(* IEC 61131-3 sources: avi-aoi-management/scripts/ai-eval/ngau-nhien/kho/st-ud7-van-hai-cuon/khung/src, 2 files *)

(* ---- ViTriVan.st ---- *)
FUNCTION ViTriVan : INT
VAR_INPUT
    CT_MO : BOOL;
    CT_DONG : BOOL;
END_VAR
    (* TODO: cài đặt theo đề bài *)
    ViTriVan := -1;
END_FUNCTION

(* ---- VanHaiCuon.st ---- *)
FUNCTION_BLOCK VanHaiCuon
VAR_INPUT
    MO : BOOL;
    DONG : BOOL;
    CT_MO : BOOL;
    CT_DONG : BOOL;
    RESET : BOOL;
    T_HANH_TRINH : TIME;
END_VAR
VAR_OUTPUT
    CUON_MO : BOOL;
    CUON_DONG : BOOL;
    TRANG_THAI : INT;
    MA_LOI : INT;
END_VAR
    (* TODO: cài đặt theo đề bài *)
    CUON_MO := FALSE;
END_FUNCTION_BLOCK
